(* IEC 61131-3 sources: kns-port-domestic/tools/inventory_tests/fixtures/lib/tests/POUs/FB_Base_Test, 1 file *)

(* ---- FB_Base_Test.decl.st ---- *)
// Назначение: набор тестов
FUNCTION_BLOCK FB_Base_Test EXTENDS coUnit.FB_TestSuite
VAR
    fbChild : FB_Child;
END_VAR
